Staubli VAL3: deleteTraj.pgx

public program deleteTraj(string x_sKey, bool& x_bToSave)
begin
  if isDefined(trajTemp:tTrajItem[x_sKey])
    delete(trajTemp:tTrajItem[x_sKey])
    //trajTemp:libSave()
  endIf
  x_bToSave=true
end
